// TIA Portal V18 export
TYPE "TaktModeZone_Input"
   STRUCT
      ModeZone_Done : Bool;
   END_STRUCT;
END_TYPE
